// Mitsubishi GX Works2 project: Practica e   PLC: FX3G

PROGRAM MAIN
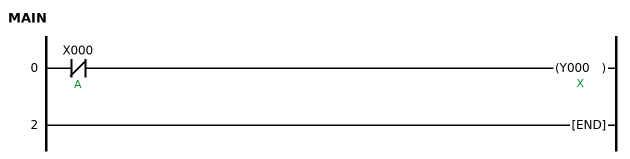
0     LDI     X000  ; A
      OUT     Y000  ; X
2     END
END_PROGRAM
